(* IEC 61131-3 sources: PLC-Static-Analysis/modules/plc-rules/src/test/resources/PLCA-Q003, 2 files *)

(* ---- compliant.st ---- *)
FUNCTION_BLOCK FB_FloatOk
VAR_INPUT
    r : REAL;
    n : INT;
END_VAR
VAR_OUTPUT
    b : BOOL;
END_VAR
VAR CONSTANT
    cA : REAL := 1.0;
    cB : REAL := 2.0;
END_VAR
b := ABS(r - 1.5) < 0.001;
b := n = 3;
b := r > 1.0;
b := cA = cB;
b := r = 0.0;
b := r <> 0;
b := r = r;
END_FUNCTION_BLOCK

(* ---- noncompliant.st ---- *)
FUNCTION_BLOCK FB_Float
VAR_INPUT
    r : REAL;
    lr : LREAL;
    n : INT;
END_VAR
VAR_OUTPUT
    b : BOOL;
END_VAR
b := r = 1.5; // PLCA-Q003
IF lr <> r THEN // PLCA-Q003
    b := FALSE;
END_IF
b := n = 0.5; // PLCA-Q003
b := r * 2.0 = INT_TO_REAL(n); // PLCA-Q003
END_FUNCTION_BLOCK
